(* IEC 61131-3 sources: TetherPLC/compat/tc2 (part 3) *)

(* ---- tc2_mc2_drive.st ---- *)
// tc2_mc2_drive.st — Tc2_MC2_Drive compatibility surface.
//
// TwinCAT's MC2 drive library addresses drives through AXIS_REF
// (here the flattened FB_MotionAxis UDINT handle, same convention
// as tc2_mc2.st).  Two transport families are covered:
//
//   CoE / OD  — CiA-402 object dictionary access through
//               FB_MotionAxis OP4/OP5 (works on both the in-process
//               tplc-motion backend and the Tether IO backend).
//               Manufacturer-specific sim objects 0x2002..0x2009
//               carry position offset, brake/park/CoE commands and
//               flying-saw characteristics (stored state, no
//               physical effect — documented).
//   SoE       — Sercos-over-EtherCAT mailbox through the builtin
//               FB_Soe (tplc-soe service, Tether IO only).  The
//               AXIS_REF handle maps to the SoE port as slave =
//               handle - 1 (MotionIoService assigns handle =
//               slave + 1).  In-process there is no SoE service,
//               so SoE FBs report bError/nErrorId = 99.
//
// NAME COLLISION NOTE: the SoE/AX5000 FB names match
// compat/tc2/tc2_drive.st (TwinCAT uses the same names in both
// libraries, differing only in the drive reference type).  This
// dialect has no library namespaces — link tc2_mc2_drive.st OR
// tc2_drive.st into a program, not both.
//
// Mapping notes (documented deviations):
//   - E_* enums (E_ParkMode, E_BrakeMode, E_PositionOffsetFeedback,
//     E_PositionOffsetMemory, E_DriveParameterNumber,
//     E_ReadWriteMode) are flattened to UDINT/INT inputs; values
//     are passed through to the backing object or ignored where
//     the sim has no equivalent.
//   - PVOID/ANY buffers (FB_CoERead/Write, FB_WriteDriveParameter)
//     are flattened to a single DINT Value; sub-index and
//     CompleteAccess are accepted but only sub-index 0 scalar
//     access is modeled.
//   - T_AmsNetID inputs are accepted for signature fidelity and
//     ignored (the axis reference already selects the drive).
//   - The 0x2002..0x2009 objects are stored command/state, not
//     physical: position offset is recorded but not applied to
//     motion, brake/park/CoE commands are recorded, saw
//     characteristics are read/write storage.
//
// SPDX-License-Identifier: Apache-2.0 OR MPL-2.0

// ---- shared helpers ------------------------------------------------
// SoE slave resolution: AXIS_REF handle -> SoE port address.
// (inlined per FB; handle = slave + 1 on the Tether IO backend)

// ================================================================== //
// §4.1 General Beckhoff
// ================================================================== //

// FB_ReadDriveParameter — read a drive parameter (OD object).
// ParameterNumber is the CiA402 object index; Mode 0 = single shot
// on Execute edge, Mode 1 = cyclic re-read while Execute is held
// (Interval is accepted; the scan rate is the cycle).
FUNCTION_BLOCK FB_ReadDriveParameter
VAR_INPUT
    Execute : BOOL;
    ParameterNumber : UDINT;
    Mode : UDINT;
    Interval : UDINT;
    Axis : UDINT;
END_VAR
VAR_OUTPUT
    Valid : BOOL;
    Value : DINT;
    Busy : BOOL;
    Done : BOOL;
    Error : BOOL;
    ErrorID : UDINT;
END_VAR
VAR
    ax : FB_MotionAxis;
    exPrev : BOOL;
    exEdge : BOOL;
END_VAR
    ax.AXIS := Axis;
    exEdge := Execute AND NOT exPrev; exPrev := Execute;
    Valid := FALSE; Busy := FALSE; Done := FALSE;
    Error := FALSE; ErrorID := 0;
    IF exEdge OR (Mode = 1 AND Execute) THEN
        ax.OP := 4;
        ax.INDEX := UDINT_TO_DINT(ParameterNumber);
        ax();
        IF ax.STATUS = 0 THEN
            Value := ax.VALUE;
            Valid := TRUE;
            IF exEdge THEN Done := TRUE; END_IF;
        ELSE
            Error := TRUE; ErrorID := ax.ERRID;
        END_IF;
    END_IF;
END_FUNCTION_BLOCK

// FB_WriteDriveParameter — write a drive parameter (OD object).
// Value is the flattened ANY buffer (single i32).
FUNCTION_BLOCK FB_WriteDriveParameter
VAR_INPUT
    Execute : BOOL;
    ParameterNumber : UDINT;
    Mode : UDINT;
    Interval : UDINT;
    Value : DINT;
    Axis : UDINT;
END_VAR
VAR_OUTPUT
    Valid : BOOL;
    Busy : BOOL;
    Done : BOOL;
    Error : BOOL;
    ErrorID : UDINT;
END_VAR
VAR
    ax : FB_MotionAxis;
    exPrev : BOOL;
    exEdge : BOOL;
END_VAR
    ax.AXIS := Axis;
    exEdge := Execute AND NOT exPrev; exPrev := Execute;
    Valid := FALSE; Busy := FALSE; Done := FALSE;
    Error := FALSE; ErrorID := 0;
    IF exEdge THEN
        ax.OP := 5;
        ax.INDEX := UDINT_TO_DINT(ParameterNumber);
        ax.VALUE := Value;
        ax();
        IF ax.STATUS = 0 THEN
            Valid := TRUE;
            Done := TRUE;
        ELSE
            Error := TRUE; ErrorID := ax.ERRID;
        END_IF;
    END_IF;
END_FUNCTION_BLOCK

// FB_SetPositionOffset — store a position offset (OD 0x2002).
// Absolute mode: offset = Position - PositionActualValue.
// Relative mode: offset accumulates (old + Position).  Feedback
// and Memory select encoder/drive/nameplate in TwinCAT; the sim
// has a single offset object, both are accepted and ignored.
FUNCTION_BLOCK FB_SetPositionOffset
VAR_INPUT
    Execute : BOOL;
    Position : LREAL;
    Relative : BOOL;
    Feedback : UDINT;
    Memory : UDINT;
    Axis : UDINT;
END_VAR
VAR_OUTPUT
    Busy : BOOL;
    Done : BOOL;
    Error : BOOL;
    ErrorID : UDINT;
END_VAR
VAR
    ax : FB_MotionAxis;
    exPrev : BOOL;
    exEdge : BOOL;
    posAct : DINT;
    offCur : DINT;
    np : DINT;
    p : DINT;
END_VAR
    ax.AXIS := Axis;
    exEdge := Execute AND NOT exPrev; exPrev := Execute;
    Busy := FALSE; Done := FALSE; Error := FALSE; ErrorID := 0;
    IF exEdge THEN
        p := LREAL_TO_DINT(Position);
        IF Relative THEN
            ax.OP := 4; ax.INDEX := 16#2002; ax();
            offCur := ax.VALUE;
            np := offCur + p;
        ELSE
            ax.OP := 4; ax.INDEX := 16#6064; ax();
            posAct := ax.VALUE;
            np := p - posAct;
        END_IF;
        ax.OP := 5; ax.INDEX := 16#2002; ax.VALUE := np; ax();
        IF ax.STATUS = 0 THEN
            Done := TRUE;
        ELSE
            Error := TRUE; ErrorID := ax.ERRID;
        END_IF;
    END_IF;
END_FUNCTION_BLOCK

// FB_DeletePositionOffset — clear the position offset (OD 0x2002).
FUNCTION_BLOCK FB_DeletePositionOffset
VAR_INPUT
    Execute : BOOL;
    Feedback : UDINT;
    Memory : UDINT;
    Axis : UDINT;
END_VAR
VAR_OUTPUT
    Busy : BOOL;
    Done : BOOL;
    Error : BOOL;
    ErrorID : UDINT;
END_VAR
VAR
    ax : FB_MotionAxis;
    exPrev : BOOL;
    exEdge : BOOL;
END_VAR
    ax.AXIS := Axis;
    exEdge := Execute AND NOT exPrev; exPrev := Execute;
    Busy := FALSE; Done := FALSE; Error := FALSE; ErrorID := 0;
    IF exEdge THEN
        ax.OP := 5; ax.INDEX := 16#2002; ax.VALUE := 0; ax();
        IF ax.STATUS = 0 THEN
            Done := TRUE;
        ELSE
            Error := TRUE; ErrorID := ax.ERRID;
        END_IF;
    END_IF;
END_FUNCTION_BLOCK

// FB_BrakeControl — brake command (OD 0x2003).  Mode is stored
// raw; the sim records the command without physical effect.
FUNCTION_BLOCK FB_BrakeControl
VAR_INPUT
    Execute : BOOL;
    Mode : UDINT;
    Axis : UDINT;
END_VAR
VAR_OUTPUT
    Busy : BOOL;
    Done : BOOL;
    Error : BOOL;
    ErrorID : UDINT;
END_VAR
VAR
    ax : FB_MotionAxis;
    exPrev : BOOL;
    exEdge : BOOL;
END_VAR
    ax.AXIS := Axis;
    exEdge := Execute AND NOT exPrev; exPrev := Execute;
    Busy := FALSE; Done := FALSE; Error := FALSE; ErrorID := 0;
    IF exEdge THEN
        ax.OP := 5; ax.INDEX := 16#2003;
        ax.VALUE := UDINT_TO_DINT(Mode); ax();
        IF ax.STATUS = 0 THEN
            Done := TRUE;
        ELSE
            Error := TRUE; ErrorID := ax.ERRID;
        END_IF;
    END_IF;
END_FUNCTION_BLOCK

// FB_ParkAxis — park/release via the SoE park mailbox (OP 7).
// Mode 0 = release, nonzero = park.  Requires the SoE backend
// (Tether IO); in-process reports bError.
FUNCTION_BLOCK FB_ParkAxis
VAR_INPUT
    Execute : BOOL;
    Mode : UDINT;
    NetId : STRING[15];
    Axis : UDINT;
END_VAR
VAR_OUTPUT
    Busy : BOOL;
    Done : BOOL;
    Error : BOOL;
    ErrorID : UDINT;
END_VAR
VAR
    raw : FB_Soe;
    exPrev : BOOL;
    exEdge : BOOL;
    slave : UDINT;
END_VAR
    exEdge := Execute AND NOT exPrev; exPrev := Execute;
    IF Axis > 0 THEN slave := Axis - 1; ELSE slave := 0; END_IF;
    Busy := FALSE; Done := FALSE; Error := FALSE; ErrorID := 0;
    IF exEdge THEN
        raw.OP := 7;
        raw.SLAVE := slave;
        IF Mode <> 0 THEN raw.VALUE := 1; ELSE raw.VALUE := 0; END_IF;
        raw();
        IF raw.STATUS < 0 THEN
            Error := TRUE; ErrorID := raw.ERRID;
        ELSE
            Done := TRUE;
        END_IF;
    END_IF;
END_FUNCTION_BLOCK

// FB_ReadDriveInfo — axis/drive info snapshot (FB_MotionAxis OP6).
FUNCTION_BLOCK FB_ReadDriveInfo
VAR_INPUT
    Execute : BOOL;
    Axis : UDINT;
END_VAR
VAR_OUTPUT
    Valid : BOOL;
    State : DINT;
    Fault : DINT;
    ModeOp : DINT;
    TargetReached : BOOL;
    PosActual : DINT;
    VelActual : DINT;
    Busy : BOOL;
    Done : BOOL;
    Error : BOOL;
    ErrorID : UDINT;
END_VAR
VAR
    ax : FB_MotionAxis;
    exPrev : BOOL;
    exEdge : BOOL;
END_VAR
    ax.AXIS := Axis;
    exEdge := Execute AND NOT exPrev; exPrev := Execute;
    Valid := FALSE; Busy := FALSE; Done := FALSE;
    Error := FALSE; ErrorID := 0;
    IF exEdge THEN
        ax.OP := 6; ax();
        IF ax.STATUS < 0 THEN
            Error := TRUE; ErrorID := ax.ERRID;
        ELSE
            Valid := TRUE;
            Done := TRUE;
            State := ax.STATUS;
            Fault := ax.FAULT;
            ModeOp := ax.MODE;
            TargetReached := (ax.TARGET_REACHED <> 0);
            PosActual := ax.POS_ACTUAL;
            VelActual := ax.VEL_ACTUAL;
        END_IF;
    END_IF;
END_FUNCTION_BLOCK

// ================================================================== //
// §4.2 General SoE
// ================================================================== //
// All SoE FBs resolve slave = Axis - 1 and drive the FB_Soe builtin.

// FB_SoERead — generic SoE element read.  Index is the SoE element
// id; the supported subset is the state-snapshot fields:
//   16#0135 -> status word (S-0-0135), 16#0267 -> password.
// Other element ids report Error (arbitrary P-0-xxxx access is not
// modeled).  Value is LREAL; u16/u32 fields are returned raw.
FUNCTION_BLOCK FB_SoERead
VAR_INPUT
    Execute : BOOL;
    Index : UDINT;
    NetId : STRING[15];
    Axis : UDINT;
END_VAR
VAR_OUTPUT
    Value : LREAL;
    Busy : BOOL;
    Done : BOOL;
    Error : BOOL;
    ErrorID : UDINT;
END_VAR
VAR
    raw : FB_Soe;
    exPrev : BOOL;
    exEdge : BOOL;
    slave : UDINT;
END_VAR
    exEdge := Execute AND NOT exPrev; exPrev := Execute;
    IF Axis > 0 THEN slave := Axis - 1; ELSE slave := 0; END_IF;
    Busy := FALSE; Done := FALSE; Error := FALSE; ErrorID := 0;
    IF exEdge THEN
        raw.OP := 1;
        raw.SLAVE := slave;
        raw();
        IF raw.STATUS < 0 THEN
            Error := TRUE; ErrorID := raw.ERRID;
        ELSE
            IF Index = 16#0135 THEN
                Value := UDINT_TO_LREAL(raw.STATUSW);
                Done := TRUE;
            ELSIF Index = 16#0267 THEN
                Value := UDINT_TO_LREAL(raw.PASSWD);
                Done := TRUE;
            ELSE
                Error := TRUE; ErrorID := 2;
            END_IF;
        END_IF;
    END_IF;
END_FUNCTION_BLOCK

// FB_SoEWrite — generic SoE element write.  Supported subset:
// Index 16#0267 -> drive password (S-0-0267).  Other ids report
// Error (arbitrary P-0-xxxx writes are not modeled).
FUNCTION_BLOCK FB_SoEWrite
VAR_INPUT
    Execute : BOOL;
    Index : UDINT;
    Value : DINT;
    NetId : STRING[15];
    Axis : UDINT;
END_VAR
VAR_OUTPUT
    Busy : BOOL;
    Done : BOOL;
    Error : BOOL;
    ErrorID : UDINT;
END_VAR
VAR
    raw : FB_Soe;
    exPrev : BOOL;
    exEdge : BOOL;
    slave : UDINT;
END_VAR
    exEdge := Execute AND NOT exPrev; exPrev := Execute;
    IF Axis > 0 THEN slave := Axis - 1; ELSE slave := 0; END_IF;
    Busy := FALSE; Done := FALSE; Error := FALSE; ErrorID := 0;
    IF exEdge THEN
        IF Index = 16#0267 THEN
            raw.OP := 2;
            raw.SLAVE := slave;
            raw.VALUE := Value;
            raw();
            IF raw.STATUS < 0 THEN
                Error := TRUE; ErrorID := raw.ERRID;
            ELSE
                Done := TRUE;
            END_IF;
        ELSE
            Error := TRUE; ErrorID := 2;
        END_IF;
    END_IF;
END_FUNCTION_BLOCK

// FB_SoESetDataAccessMode — SoE parameter access mode.  The sim
// mailbox always uses parallel access; the FB accepts the request
// and completes (documented no-op).
FUNCTION_BLOCK FB_SoESetDataAccessMode
VAR_INPUT
    Execute : BOOL;
    Mode : UDINT;
    Axis : UDINT;
END_VAR
VAR_OUTPUT
    Busy : BOOL;
    Done : BOOL;
    Error : BOOL;
    ErrorID : UDINT;
END_VAR
VAR
    exPrev : BOOL;
    exEdge : BOOL;
END_VAR
    exEdge := Execute AND NOT exPrev; exPrev := Execute;
    Busy := FALSE; Done := FALSE; Error := FALSE; ErrorID := 0;
    IF exEdge THEN
        Done := TRUE;
    END_IF;
END_FUNCTION_BLOCK

// ---- command FBs ----------------------------------------------------

// FB_SoEReset — S-0-0099 drive reset.
FUNCTION_BLOCK FB_SoEReset
VAR_INPUT
    Execute : BOOL;
    NetId : STRING[15];
    Axis : UDINT;
END_VAR
VAR_OUTPUT
    Busy : BOOL;
    Done : BOOL;
    Error : BOOL;
    ErrorID : UDINT;
END_VAR
VAR
    raw : FB_Soe;
    exPrev : BOOL;
    exEdge : BOOL;
    slave : UDINT;
END_VAR
    exEdge := Execute AND NOT exPrev; exPrev := Execute;
    IF Axis > 0 THEN slave := Axis - 1; ELSE slave := 0; END_IF;
    Busy := FALSE; Done := FALSE; Error := FALSE; ErrorID := 0;
    IF exEdge THEN
        raw.OP := 5;
        raw.SLAVE := slave;
        raw();
        IF raw.STATUS < 0 THEN
            Error := TRUE; ErrorID := raw.ERRID;
        ELSE
            Done := TRUE;
        END_IF;
    END_IF;
END_FUNCTION_BLOCK

// FB_SoEWritePassword — S-0-0267 drive password.
FUNCTION_BLOCK FB_SoEWritePassword
VAR_INPUT
    Execute : BOOL;
    Password : UDINT;
    NetId : STRING[15];
    Axis : UDINT;
END_VAR
VAR_OUTPUT
    Busy : BOOL;
    Done : BOOL;
    Error : BOOL;
    ErrorID : UDINT;
END_VAR
VAR
    raw : FB_Soe;
    exPrev : BOOL;
    exEdge : BOOL;
    slave : UDINT;
END_VAR
    exEdge := Execute AND NOT exPrev; exPrev := Execute;
    IF Axis > 0 THEN slave := Axis - 1; ELSE slave := 0; END_IF;
    Busy := FALSE; Done := FALSE; Error := FALSE; ErrorID := 0;
    IF exEdge THEN
        raw.OP := 2;
        raw.SLAVE := slave;
        raw.VALUE := UDINT_TO_DINT(Password);
        raw();
        IF raw.STATUS < 0 THEN
            Error := TRUE; ErrorID := raw.ERRID;
        ELSE
            Done := TRUE;
        END_IF;
    END_IF;
END_FUNCTION_BLOCK

// FB_SoEExecuteCommand — execute an SoE command id.
FUNCTION_BLOCK FB_SoEExecuteCommand
VAR_INPUT
    Execute : BOOL;
    CommandId : UDINT;
    NetId : STRING[15];
    Axis : UDINT;
END_VAR
VAR_OUTPUT
    Busy : BOOL;
    Done : BOOL;
    Error : BOOL;
    ErrorID : UDINT;
END_VAR
VAR
    raw : FB_Soe;
    exPrev : BOOL;
    exEdge : BOOL;
    slave : UDINT;
END_VAR
    exEdge := Execute AND NOT exPrev; exPrev := Execute;
    IF Axis > 0 THEN slave := Axis - 1; ELSE slave := 0; END_IF;
    Busy := FALSE; Done := FALSE; Error := FALSE; ErrorID := 0;
    IF exEdge THEN
        raw.OP := 4;
        raw.SLAVE := slave;
        raw.VALUE := UDINT_TO_DINT(CommandId);
        raw();
        IF raw.STATUS < 0 THEN
            Error := TRUE; ErrorID := raw.ERRID;
        ELSE
            Done := TRUE;
        END_IF;
    END_IF;
END_FUNCTION_BLOCK

// FB_SoEWriteCommandControl — command control word.
FUNCTION_BLOCK FB_SoEWriteCommandControl
VAR_INPUT
    Execute : BOOL;
    CommandControl : UDINT;
    NetId : STRING[15];
    Axis : UDINT;
END_VAR
VAR_OUTPUT
    Busy : BOOL;
    Done : BOOL;
    Error : BOOL;
    ErrorID : UDINT;
END_VAR
VAR
    raw : FB_Soe;
    exPrev : BOOL;
    exEdge : BOOL;
    slave : UDINT;
END_VAR
    exEdge := Execute AND NOT exPrev; exPrev := Execute;
    IF Axis > 0 THEN slave := Axis - 1; ELSE slave := 0; END_IF;
    Busy := FALSE; Done := FALSE; Error := FALSE; ErrorID := 0;
    IF exEdge THEN
        raw.OP := 3;
        raw.SLAVE := slave;
        raw.VALUE := UDINT_TO_DINT(CommandControl);
        raw();
        IF raw.STATUS < 0 THEN
            Error := TRUE; ErrorID := raw.ERRID;
        ELSE
            Done := TRUE;
        END_IF;
    END_IF;
END_FUNCTION_BLOCK

// FB_SoEReadCommandState — SoE command state
// (0 idle, 1 running, 2 done, 3 error).
FUNCTION_BLOCK FB_SoEReadCommandState
VAR_INPUT
    Execute : BOOL;
    NetId : STRING[15];
    Axis : UDINT;
END_VAR
VAR_OUTPUT
    CommandState : UDINT;
    Busy : BOOL;
    Done : BOOL;
    Error : BOOL;
    ErrorID : UDINT;
END_VAR
VAR
    raw : FB_Soe;
    exPrev : BOOL;
    exEdge : BOOL;
    slave : UDINT;
END_VAR
    exEdge := Execute AND NOT exPrev; exPrev := Execute;
    IF Axis > 0 THEN slave := Axis - 1; ELSE slave := 0; END_IF;
    Busy := FALSE; Done := FALSE; Error := FALSE; ErrorID := 0;
    IF exEdge THEN
        raw.OP := 1;
        raw.SLAVE := slave;
        raw();
        IF raw.STATUS < 0 THEN
            Error := TRUE; ErrorID := raw.ERRID;
        ELSE
            CommandState := raw.CMDSTATE;
            Done := TRUE;
        END_IF;
    END_IF;
END_FUNCTION_BLOCK

// ---- diagnostics FBs -------------------------------------------------

// FB_SoEReadDiagMessage — S-0-0095 diagnosis message.
FUNCTION_BLOCK FB_SoEReadDiagMessage
VAR_INPUT
    Execute : BOOL;
    NetId : STRING[15];
    Axis : UDINT;
END_VAR
VAR_OUTPUT
    DiagMessage : STRING[63];
    Busy : BOOL;
    Done : BOOL;
    Error : BOOL;
    ErrorID : UDINT;
END_VAR
VAR
    raw : FB_Soe;
    exPrev : BOOL;
    exEdge : BOOL;
    slave : UDINT;
END_VAR
    exEdge := Execute AND NOT exPrev; exPrev := Execute;
    IF Axis > 0 THEN slave := Axis - 1; ELSE slave := 0; END_IF;
    Busy := FALSE; Done := FALSE; Error := FALSE; ErrorID := 0;
    IF exEdge THEN
        raw.OP := 1;
        raw.SLAVE := slave;
        raw();
        IF raw.STATUS < 0 THEN
            Error := TRUE; ErrorID := raw.ERRID;
        ELSE
            DiagMessage := raw.DIAGMSG;
            Done := TRUE;
        END_IF;
    END_IF;
END_FUNCTION_BLOCK

// FB_SoEReadDiagNumber — diagnosis number.
FUNCTION_BLOCK FB_SoEReadDiagNumber
VAR_INPUT
    Execute : BOOL;
    NetId : STRING[15];
    Axis : UDINT;
END_VAR
VAR_OUTPUT
    DiagNumber : UDINT;
    Busy : BOOL;
    Done : BOOL;
    Error : BOOL;
    ErrorID : UDINT;
END_VAR
VAR
    raw : FB_Soe;
    exPrev : BOOL;
    exEdge : BOOL;
    slave : UDINT;
END_VAR
    exEdge := Execute AND NOT exPrev; exPrev := Execute;
    IF Axis > 0 THEN slave := Axis - 1; ELSE slave := 0; END_IF;
    Busy := FALSE; Done := FALSE; Error := FALSE; ErrorID := 0;
    IF exEdge THEN
        raw.OP := 1;
        raw.SLAVE := slave;
        raw();
        IF raw.STATUS < 0 THEN
            Error := TRUE; ErrorID := raw.ERRID;
        ELSE
            DiagNumber := raw.DIAGNUM;
            Done := TRUE;
        END_IF;
    END_IF;
END_FUNCTION_BLOCK

// FB_SoEReadDiagNumberList — diagnosis number list (flattened:
// DiagCount + DiagList internal array).
FUNCTION_BLOCK FB_SoEReadDiagNumberList
VAR_INPUT
    Execute : BOOL;
    NetId : STRING[15];
    Axis : UDINT;
END_VAR
VAR_OUTPUT
    DiagCount : UDINT;
    Busy : BOOL;
    Done : BOOL;
    Error : BOOL;
    ErrorID : UDINT;
END_VAR
VAR
    raw : FB_Soe;
    exPrev : BOOL;
    exEdge : BOOL;
    slave : UDINT;
    i : UDINT;
    DiagList : ARRAY[0..7] OF UDINT;
END_VAR
    exEdge := Execute AND NOT exPrev; exPrev := Execute;
    IF Axis > 0 THEN slave := Axis - 1; ELSE slave := 0; END_IF;
    Busy := FALSE; Done := FALSE; Error := FALSE; ErrorID := 0;
    IF exEdge THEN
        raw.OP := 1;
        raw.SLAVE := slave;
        raw();
        IF raw.STATUS < 0 THEN
            Error := TRUE; ErrorID := raw.ERRID;
        ELSE
            DiagCount := raw.DIAGCOUNT;
            FOR i := 0 TO 7 DO
                DiagList[i] := raw.DIAGLIST[i];
            END_FOR;
            Done := TRUE;
        END_IF;
    END_IF;
END_FUNCTION_BLOCK

// FB_SoEReadClassXDiag — class-X diagnosis.
FUNCTION_BLOCK FB_SoEReadClassXDiag
VAR_INPUT
    Execute : BOOL;
    NetId : STRING[15];
    Axis : UDINT;
END_VAR
VAR_OUTPUT
    ClassXDiag : UDINT;
    Busy : BOOL;
    Done : BOOL;
    Error : BOOL;
    ErrorID : UDINT;
END_VAR
VAR
    raw : FB_Soe;
    exPrev : BOOL;
    exEdge : BOOL;
    slave : UDINT;
END_VAR
    exEdge := Execute AND NOT exPrev; exPrev := Execute;
    IF Axis > 0 THEN slave := Axis - 1; ELSE slave := 0; END_IF;
    Busy := FALSE; Done := FALSE; Error := FALSE; ErrorID := 0;
    IF exEdge THEN
        raw.OP := 1;
        raw.SLAVE := slave;
        raw();
        IF raw.STATUS < 0 THEN
            Error := TRUE; ErrorID := raw.ERRID;
        ELSE
            ClassXDiag := raw.CLASSX;
            Done := TRUE;
        END_IF;
    END_IF;
END_FUNCTION_BLOCK

// ---- current-value readers -------------------------------------------

FUNCTION_BLOCK FB_SoEReadAmplifierTemperature
VAR_INPUT
    Execute : BOOL;
    NetId : STRING[15];
    Axis : UDINT;
END_VAR
VAR_OUTPUT
    Value : LREAL;
    Busy : BOOL;
    Done : BOOL;
    Error : BOOL;
    ErrorID : UDINT;
END_VAR
VAR
    raw : FB_Soe;
    exPrev : BOOL;
    exEdge : BOOL;
    slave : UDINT;
END_VAR
    exEdge := Execute AND NOT exPrev; exPrev := Execute;
    IF Axis > 0 THEN slave := Axis - 1; ELSE slave := 0; END_IF;
    Busy := FALSE; Done := FALSE; Error := FALSE; ErrorID := 0;
    IF exEdge THEN
        raw.OP := 1;
        raw.SLAVE := slave;
        raw();
        IF raw.STATUS < 0 THEN
            Error := TRUE; ErrorID := raw.ERRID;
        ELSE
            Value := raw.AMPTEMP;
            Done := TRUE;
        END_IF;
    END_IF;
END_FUNCTION_BLOCK

FUNCTION_BLOCK FB_SoEReadMotorTemperature
VAR_INPUT
    Execute : BOOL;
    NetId : STRING[15];
    Axis : UDINT;
END_VAR
VAR_OUTPUT
    Value : LREAL;
    Busy : BOOL;
    Done : BOOL;
    Error : BOOL;
    ErrorID : UDINT;
END_VAR
VAR
    raw : FB_Soe;
    exPrev : BOOL;
    exEdge : BOOL;
    slave : UDINT;
END_VAR
    exEdge := Execute AND NOT exPrev; exPrev := Execute;
    IF Axis > 0 THEN slave := Axis - 1; ELSE slave := 0; END_IF;
    Busy := FALSE; Done := FALSE; Error := FALSE; ErrorID := 0;
    IF exEdge THEN
        raw.OP := 1;
        raw.SLAVE := slave;
        raw();
        IF raw.STATUS < 0 THEN
            Error := TRUE; ErrorID := raw.ERRID;
        ELSE
            Value := raw.MTEMPT;
            Done := TRUE;
        END_IF;
    END_IF;
END_FUNCTION_BLOCK

FUNCTION_BLOCK FB_SoEReadDcBusVoltage
VAR_INPUT
    Execute : BOOL;
    NetId : STRING[15];
    Axis : UDINT;
END_VAR
VAR_OUTPUT
    Value : LREAL;
    Busy : BOOL;
    Done : BOOL;
    Error : BOOL;
    ErrorID : UDINT;
END_VAR
VAR
    raw : FB_Soe;
    exPrev : BOOL;
    exEdge : BOOL;
    slave : UDINT;
END_VAR
    exEdge := Execute AND NOT exPrev; exPrev := Execute;
    IF Axis > 0 THEN slave := Axis - 1; ELSE slave := 0; END_IF;
    Busy := FALSE; Done := FALSE; Error := FALSE; ErrorID := 0;
    IF exEdge THEN
        raw.OP := 1;
        raw.SLAVE := slave;
        raw();
        IF raw.STATUS < 0 THEN
            Error := TRUE; ErrorID := raw.ERRID;
        ELSE
            Value := raw.DCVOLT;
            Done := TRUE;
        END_IF;
    END_IF;
END_FUNCTION_BLOCK

FUNCTION_BLOCK FB_SoEReadDcBusCurrent
VAR_INPUT
    Execute : BOOL;
    NetId : STRING[15];
    Axis : UDINT;
END_VAR
VAR_OUTPUT
    Value : LREAL;
    Busy : BOOL;
    Done : BOOL;
    Error : BOOL;
    ErrorID : UDINT;
END_VAR
VAR
    raw : FB_Soe;
    exPrev : BOOL;
    exEdge : BOOL;
    slave : UDINT;
END_VAR
    exEdge := Execute AND NOT exPrev; exPrev := Execute;
    IF Axis > 0 THEN slave := Axis - 1; ELSE slave := 0; END_IF;
    Busy := FALSE; Done := FALSE; Error := FALSE; ErrorID := 0;
    IF exEdge THEN
        raw.OP := 1;
        raw.SLAVE := slave;
        raw();
        IF raw.STATUS < 0 THEN
            Error := TRUE; ErrorID := raw.ERRID;
        ELSE
            Value := raw.DCCURR;
            Done := TRUE;
        END_IF;
    END_IF;
END_FUNCTION_BLOCK

// ================================================================== //
// §4.3 General CoE — SDO object access via FB_MotionAxis OP4/OP5.
// Index/SubIndex select the object; SubIndex and CompleteAccess are
// accepted but only sub-index 0 scalar access is modeled.  Value is
// the flattened PVOID buffer (single i32).
// ================================================================== //

// FB_CoERead — CoE SDO upload.
FUNCTION_BLOCK FB_CoERead
VAR_INPUT
    Execute : BOOL;
    Index : UDINT;
    SubIndex : UDINT;
    CompleteAccess : BOOL;
    NetId : STRING[15];
    Axis : UDINT;
END_VAR
VAR_OUTPUT
    Value : DINT;
    Busy : BOOL;
    Done : BOOL;
    Error : BOOL;
    ErrorID : UDINT;
END_VAR
VAR
    ax : FB_MotionAxis;
    exPrev : BOOL;
    exEdge : BOOL;
END_VAR
    ax.AXIS := Axis;
    exEdge := Execute AND NOT exPrev; exPrev := Execute;
    Busy := FALSE; Done := FALSE; Error := FALSE; ErrorID := 0;
    IF exEdge THEN
        IF SubIndex <> 0 THEN
            Error := TRUE; ErrorID := 2;   // sub-index unsupported
        ELSE
            ax.OP := 4;
            ax.INDEX := UDINT_TO_DINT(Index);
            ax();
            IF ax.STATUS = 0 THEN
                Value := ax.VALUE;
                Done := TRUE;
            ELSE
                Error := TRUE; ErrorID := ax.ERRID;
            END_IF;
        END_IF;
    END_IF;
END_FUNCTION_BLOCK

// FB_CoEWrite — CoE SDO download.
FUNCTION_BLOCK FB_CoEWrite
VAR_INPUT
    Execute : BOOL;
    Index : UDINT;
    SubIndex : UDINT;
    Value : DINT;
    CompleteAccess : BOOL;
    NetId : STRING[15];
    Axis : UDINT;
END_VAR
VAR_OUTPUT
    Busy : BOOL;
    Done : BOOL;
    Error : BOOL;
    ErrorID : UDINT;
END_VAR
VAR
    ax : FB_MotionAxis;
    exPrev : BOOL;
    exEdge : BOOL;
END_VAR
    ax.AXIS := Axis;
    exEdge := Execute AND NOT exPrev; exPrev := Execute;
    Busy := FALSE; Done := FALSE; Error := FALSE; ErrorID := 0;
    IF exEdge THEN
        IF SubIndex <> 0 THEN
            Error := TRUE; ErrorID := 2;
        ELSE
            ax.OP := 5;
            ax.INDEX := UDINT_TO_DINT(Index);
            ax.VALUE := Value;
            ax();
            IF ax.STATUS = 0 THEN
                Done := TRUE;
            ELSE
                Error := TRUE; ErrorID := ax.ERRID;
            END_IF;
        END_IF;
    END_IF;
END_FUNCTION_BLOCK

// FB_CoEExecuteCommand — execute a CoE drive command (OD 0x2005).
// Command is the flattened command id; the sim records it.
FUNCTION_BLOCK FB_CoEExecuteCommand
VAR_INPUT
    Execute : BOOL;
    Command : UDINT;
    NetId : STRING[15];
    Axis : UDINT;
END_VAR
VAR_OUTPUT
    Busy : BOOL;
    Done : BOOL;
    Error : BOOL;
    ErrorID : UDINT;
END_VAR
VAR
    ax : FB_MotionAxis;
    exPrev : BOOL;
    exEdge : BOOL;
END_VAR
    ax.AXIS := Axis;
    exEdge := Execute AND NOT exPrev; exPrev := Execute;
    Busy := FALSE; Done := FALSE; Error := FALSE; ErrorID := 0;
    IF exEdge THEN
        ax.OP := 5; ax.INDEX := 16#2005;
        ax.VALUE := UDINT_TO_DINT(Command); ax();
        IF ax.STATUS = 0 THEN
            Done := TRUE;
        ELSE
            Error := TRUE; ErrorID := ax.ERRID;
        END_IF;
    END_IF;
END_FUNCTION_BLOCK

// ================================================================== //
// §4.4 AX5000 SoE — same SoE mailbox surface as the general blocks,
// AX5000-specific objects (mains voltage, motor ctrl word, firmware,
// park, position offset).
// ================================================================== //

// FB_SoEAX5000ReadActMainVoltage — P-0-0200 peak mains voltage.
FUNCTION_BLOCK FB_SoEAX5000ReadActMainVoltage
VAR_INPUT
    Execute : BOOL;
    NetId : STRING[15];
    Axis : UDINT;
END_VAR
VAR_OUTPUT
    Voltage : LREAL;
    Busy : BOOL;
    Done : BOOL;
    Error : BOOL;
    ErrorID : UDINT;
END_VAR
VAR
    raw : FB_Soe;
    exPrev : BOOL;
    exEdge : BOOL;
    slave : UDINT;
END_VAR
    exEdge := Execute AND NOT exPrev; exPrev := Execute;
    IF Axis > 0 THEN slave := Axis - 1; ELSE slave := 0; END_IF;
    Busy := FALSE; Done := FALSE; Error := FALSE; ErrorID := 0;
    IF exEdge THEN
        raw.OP := 1;
        raw.SLAVE := slave;
        raw();
        IF raw.STATUS < 0 THEN
            Error := TRUE; ErrorID := raw.ERRID;
        ELSE
            Voltage := raw.AXMAINS;
            Done := TRUE;
        END_IF;
    END_IF;
END_FUNCTION_BLOCK

// FB_SoEAX5000SetMotorCtrlWord — motor control word (mailbox OP6).
// bForceUnlock accepted for signature compatibility.
FUNCTION_BLOCK FB_SoEAX5000SetMotorCtrlWord
VAR_INPUT
    Execute : BOOL;
    MotorCtrlWord : UDINT;
    bForceUnlock : BOOL;
    NetId : STRING[15];
    Axis : UDINT;
END_VAR
VAR_OUTPUT
    Busy : BOOL;
    Done : BOOL;
    Error : BOOL;
    ErrorID : UDINT;
END_VAR
VAR
    raw : FB_Soe;
    exPrev : BOOL;
    exEdge : BOOL;
    slave : UDINT;
END_VAR
    exEdge := Execute AND NOT exPrev; exPrev := Execute;
    IF Axis > 0 THEN slave := Axis - 1; ELSE slave := 0; END_IF;
    Busy := FALSE; Done := FALSE; Error := FALSE; ErrorID := 0;
    IF exEdge THEN
        raw.OP := 6;
        raw.SLAVE := slave;
        raw.VALUE := UDINT_TO_DINT(MotorCtrlWord);
        raw();
        IF raw.STATUS < 0 THEN
            Error := TRUE; ErrorID := raw.ERRID;
        ELSE
            Done := TRUE;
        END_IF;
    END_IF;
END_FUNCTION_BLOCK

// FB_SoEAX5000FirmwareUpdate — reports simulated firmware
// revision/build; no firmware pool or flashing is simulated.
FUNCTION_BLOCK FB_SoEAX5000FirmwareUpdate
VAR_INPUT
    Execute : BOOL;
    NetId : STRING[15];
    Axis : UDINT;
END_VAR
VAR_OUTPUT
    FirmwareRevision : UDINT;
    FirmwareBuild : UDINT;
    Busy : BOOL;
    Done : BOOL;
    Error : BOOL;
    ErrorID : UDINT;
END_VAR
VAR
    raw : FB_Soe;
    exPrev : BOOL;
    exEdge : BOOL;
    slave : UDINT;
END_VAR
    exEdge := Execute AND NOT exPrev; exPrev := Execute;
    IF Axis > 0 THEN slave := Axis - 1; ELSE slave := 0; END_IF;
    Busy := FALSE; Done := FALSE; Error := FALSE; ErrorID := 0;
    IF exEdge THEN
        raw.OP := 1;
        raw.SLAVE := slave;
        raw();
        IF raw.STATUS < 0 THEN
            Error := TRUE; ErrorID := raw.ERRID;
        ELSE
            FirmwareRevision := raw.AXFWREV;
            FirmwareBuild := raw.AXFWBUILD;
            Done := TRUE;
        END_IF;
    END_IF;
END_FUNCTION_BLOCK

// FB_SoEAX5000SetPositionOffset — AX5000 position offset (OD 0x2002).
FUNCTION_BLOCK FB_SoEAX5000SetPositionOffset
VAR_INPUT
    Execute : BOOL;
    Position : LREAL;
    Relative : BOOL;
    Feedback : UDINT;
    Memory : UDINT;
    NetId : STRING[15];
    Axis : UDINT;
END_VAR
VAR_OUTPUT
    Busy : BOOL;
    Done : BOOL;
    Error : BOOL;
    ErrorID : UDINT;
END_VAR
VAR
    ax : FB_MotionAxis;
    exPrev : BOOL;
    exEdge : BOOL;
    posAct : DINT;
    np : DINT;
    p : DINT;
END_VAR
    ax.AXIS := Axis;
    exEdge := Execute AND NOT exPrev; exPrev := Execute;
    Busy := FALSE; Done := FALSE; Error := FALSE; ErrorID := 0;
    IF exEdge THEN
        p := LREAL_TO_DINT(Position);
        IF Relative THEN
            np := p;                    // relative: offset delta
        ELSE
            ax.OP := 4; ax.INDEX := 16#6064; ax();
            posAct := ax.VALUE;
            np := p - posAct;
        END_IF;
        ax.OP := 5; ax.INDEX := 16#2002; ax.VALUE := np; ax();
        IF ax.STATUS = 0 THEN
            Done := TRUE;
        ELSE
            Error := TRUE; ErrorID := ax.ERRID;
        END_IF;
    END_IF;
END_FUNCTION_BLOCK

// FB_SoEAX5000DeletePositionOffset — clear AX5000 position offset.
FUNCTION_BLOCK FB_SoEAX5000DeletePositionOffset
VAR_INPUT
    Execute : BOOL;
    Feedback : UDINT;
    Memory : UDINT;
    NetId : STRING[15];
    Axis : UDINT;
END_VAR
VAR_OUTPUT
    Busy : BOOL;
    Done : BOOL;
    Error : BOOL;
    ErrorID : UDINT;
END_VAR
VAR
    ax : FB_MotionAxis;
    exPrev : BOOL;
    exEdge : BOOL;
END_VAR
    ax.AXIS := Axis;
    exEdge := Execute AND NOT exPrev; exPrev := Execute;
    Busy := FALSE; Done := FALSE; Error := FALSE; ErrorID := 0;
    IF exEdge THEN
        ax.OP := 5; ax.INDEX := 16#2002; ax.VALUE := 0; ax();
        IF ax.STATUS = 0 THEN
            Done := TRUE;
        ELSE
            Error := TRUE; ErrorID := ax.ERRID;
        END_IF;
    END_IF;
END_FUNCTION_BLOCK

// FB_SoEAX5000ParkAxis — park/unpark via SoE mailbox (OP 7).
FUNCTION_BLOCK FB_SoEAX5000ParkAxis
VAR_INPUT
    Execute : BOOL;
    Mode : UDINT;
    NetId : STRING[15];
    Axis : UDINT;
END_VAR
VAR_OUTPUT
    Busy : BOOL;
    Done : BOOL;
    Error : BOOL;
    ErrorID : UDINT;
END_VAR
VAR
    raw : FB_Soe;
    exPrev : BOOL;
    exEdge : BOOL;
    slave : UDINT;
END_VAR
    exEdge := Execute AND NOT exPrev; exPrev := Execute;
    IF Axis > 0 THEN slave := Axis - 1; ELSE slave := 0; END_IF;
    Busy := FALSE; Done := FALSE; Error := FALSE; ErrorID := 0;
    IF exEdge THEN
        raw.OP := 7;
        raw.SLAVE := slave;
        IF Mode <> 0 THEN raw.VALUE := 1; ELSE raw.VALUE := 0; END_IF;
        raw();
        IF raw.STATUS < 0 THEN
            Error := TRUE; ErrorID := raw.ERRID;
        ELSE
            Done := TRUE;
        END_IF;
    END_IF;
END_FUNCTION_BLOCK

// ================================================================== //
// §4.5 AX8000 CoE — brake/park/offset over OD objects 0x2002-0x2004.
// ================================================================== //

// FB_CoEAX8000BrakeControl — AX8000 brake (OD 0x2003).
FUNCTION_BLOCK FB_CoEAX8000BrakeControl
VAR_INPUT
    Execute : BOOL;
    Mode : UDINT;
    NetId : STRING[15];
    Axis : UDINT;
END_VAR
VAR_OUTPUT
    Busy : BOOL;
    Done : BOOL;
    Error : BOOL;
    ErrorID : UDINT;
END_VAR
VAR
    ax : FB_MotionAxis;
    exPrev : BOOL;
    exEdge : BOOL;
END_VAR
    ax.AXIS := Axis;
    exEdge := Execute AND NOT exPrev; exPrev := Execute;
    Busy := FALSE; Done := FALSE; Error := FALSE; ErrorID := 0;
    IF exEdge THEN
        ax.OP := 5; ax.INDEX := 16#2003;
        ax.VALUE := UDINT_TO_DINT(Mode); ax();
        IF ax.STATUS = 0 THEN
            Done := TRUE;
        ELSE
            Error := TRUE; ErrorID := ax.ERRID;
        END_IF;
    END_IF;
END_FUNCTION_BLOCK

// FB_CoEAX8000BrakeTest — brake test: writes the test command and
// reports Succeeded (the sim has no torque verification; the test
// always succeeds once the command is accepted — documented).
FUNCTION_BLOCK FB_CoEAX8000BrakeTest
VAR_INPUT
    Execute : BOOL;
    NetId : STRING[15];
    Axis : UDINT;
END_VAR
VAR_OUTPUT
    Succeeded : BOOL;
    Busy : BOOL;
    Done : BOOL;
    Error : BOOL;
    ErrorID : UDINT;
END_VAR
VAR
    ax : FB_MotionAxis;
    exPrev : BOOL;
    exEdge : BOOL;
END_VAR
    ax.AXIS := Axis;
    exEdge := Execute AND NOT exPrev; exPrev := Execute;
    Busy := FALSE; Done := FALSE; Error := FALSE; ErrorID := 0;
    Succeeded := FALSE;
    IF exEdge THEN
        ax.OP := 5; ax.INDEX := 16#2003; ax.VALUE := 2; ax();
        IF ax.STATUS = 0 THEN
            Done := TRUE;
            Succeeded := TRUE;
        ELSE
            Error := TRUE; ErrorID := ax.ERRID;
        END_IF;
    END_IF;
END_FUNCTION_BLOCK

// FB_CoEAX8000SetPositionOffset — AX8000 position offset (0x2002).
FUNCTION_BLOCK FB_CoEAX8000SetPositionOffset
VAR_INPUT
    Execute : BOOL;
    Position : LREAL;
    Relative : BOOL;
    Feedback : UDINT;
    Memory : UDINT;
    NetId : STRING[15];
    Axis : UDINT;
END_VAR
VAR_OUTPUT
    Busy : BOOL;
    Done : BOOL;
    Error : BOOL;
    ErrorID : UDINT;
END_VAR
VAR
    ax : FB_MotionAxis;
    exPrev : BOOL;
    exEdge : BOOL;
    posAct : DINT;
    np : DINT;
    p : DINT;
END_VAR
    ax.AXIS := Axis;
    exEdge := Execute AND NOT exPrev; exPrev := Execute;
    Busy := FALSE; Done := FALSE; Error := FALSE; ErrorID := 0;
    IF exEdge THEN
        p := LREAL_TO_DINT(Position);
        IF Relative THEN
            np := p;
        ELSE
            ax.OP := 4; ax.INDEX := 16#6064; ax();
            posAct := ax.VALUE;
            np := p - posAct;
        END_IF;
        ax.OP := 5; ax.INDEX := 16#2002; ax.VALUE := np; ax();
        IF ax.STATUS = 0 THEN
            Done := TRUE;
        ELSE
            Error := TRUE; ErrorID := ax.ERRID;
        END_IF;
    END_IF;
END_FUNCTION_BLOCK

// FB_CoEAX8000DeletePositionOffset — clear AX8000 offset (0x2002).
FUNCTION_BLOCK FB_CoEAX8000DeletePositionOffset
VAR_INPUT
    Execute : BOOL;
    Position : LREAL;
    Relative : BOOL;
    Feedback : UDINT;
    Memory : UDINT;
    NetId : STRING[15];
    Axis : UDINT;
END_VAR
VAR_OUTPUT
    Busy : BOOL;
    Done : BOOL;
    Error : BOOL;
    ErrorID : UDINT;
END_VAR
VAR
    ax : FB_MotionAxis;
    exPrev : BOOL;
    exEdge : BOOL;
END_VAR
    ax.AXIS := Axis;
    exEdge := Execute AND NOT exPrev; exPrev := Execute;
    Busy := FALSE; Done := FALSE; Error := FALSE; ErrorID := 0;
    IF exEdge THEN
        ax.OP := 5; ax.INDEX := 16#2002; ax.VALUE := 0; ax();
        IF ax.STATUS = 0 THEN
            Done := TRUE;
        ELSE
            Error := TRUE; ErrorID := ax.ERRID;
        END_IF;
    END_IF;
END_FUNCTION_BLOCK

// FB_CoEAX8000ParkAxis — AX8000 park via CoE object 0x2004.
FUNCTION_BLOCK FB_CoEAX8000ParkAxis
VAR_INPUT
    Execute : BOOL;
    Mode : UDINT;
    NetId : STRING[15];
    Axis : UDINT;
END_VAR
VAR_OUTPUT
    Busy : BOOL;
    Done : BOOL;
    Error : BOOL;
    ErrorID : UDINT;
END_VAR
VAR
    ax : FB_MotionAxis;
    exPrev : BOOL;
    exEdge : BOOL;
END_VAR
    ax.AXIS := Axis;
    exEdge := Execute AND NOT exPrev; exPrev := Execute;
    Busy := FALSE; Done := FALSE; Error := FALSE; ErrorID := 0;
    IF exEdge THEN
        ax.OP := 5; ax.INDEX := 16#2004;
        IF Mode <> 0 THEN ax.VALUE := 1; ELSE ax.VALUE := 0; END_IF;
        ax();
        IF ax.STATUS = 0 THEN
            Done := TRUE;
        ELSE
            Error := TRUE; ErrorID := ax.ERRID;
        END_IF;
    END_IF;
END_FUNCTION_BLOCK

// ================================================================== //
// §4.6 EL72xx CoE — brake/offset over the same OD objects.
// ================================================================== //

// FB_CoEEL72xxBrakeControl — EL72xx brake (OD 0x2003).
FUNCTION_BLOCK FB_CoEEL72xxBrakeControl
VAR_INPUT
    Execute : BOOL;
    Mode : UDINT;
    Axis : UDINT;
END_VAR
VAR_OUTPUT
    Busy : BOOL;
    Done : BOOL;
    Error : BOOL;
    ErrorID : UDINT;
END_VAR
VAR
    ax : FB_MotionAxis;
    exPrev : BOOL;
    exEdge : BOOL;
END_VAR
    ax.AXIS := Axis;
    exEdge := Execute AND NOT exPrev; exPrev := Execute;
    Busy := FALSE; Done := FALSE; Error := FALSE; ErrorID := 0;
    IF exEdge THEN
        ax.OP := 5; ax.INDEX := 16#2003;
        ax.VALUE := UDINT_TO_DINT(Mode); ax();
        IF ax.STATUS = 0 THEN
            Done := TRUE;
        ELSE
            Error := TRUE; ErrorID := ax.ERRID;
        END_IF;
    END_IF;
END_FUNCTION_BLOCK

// FB_CoEEL72xxSetPositionOffset — EL72xx offset (0x2002).
FUNCTION_BLOCK FB_CoEEL72xxSetPositionOffset
VAR_INPUT
    Execute : BOOL;
    Position : LREAL;
    Relative : BOOL;
    Feedback : UDINT;
    Memory : UDINT;
    Axis : UDINT;
END_VAR
VAR_OUTPUT
    Busy : BOOL;
    Done : BOOL;
    Error : BOOL;
    ErrorID : UDINT;
END_VAR
VAR
    ax : FB_MotionAxis;
    exPrev : BOOL;
    exEdge : BOOL;
    posAct : DINT;
    np : DINT;
    p : DINT;
END_VAR
    ax.AXIS := Axis;
    exEdge := Execute AND NOT exPrev; exPrev := Execute;
    Busy := FALSE; Done := FALSE; Error := FALSE; ErrorID := 0;
    IF exEdge THEN
        p := LREAL_TO_DINT(Position);
        IF Relative THEN
            np := p;
        ELSE
            ax.OP := 4; ax.INDEX := 16#6064; ax();
            posAct := ax.VALUE;
            np := p - posAct;
        END_IF;
        ax.OP := 5; ax.INDEX := 16#2002; ax.VALUE := np; ax();
        IF ax.STATUS = 0 THEN
            Done := TRUE;
        ELSE
            Error := TRUE; ErrorID := ax.ERRID;
        END_IF;
    END_IF;
END_FUNCTION_BLOCK

// FB_CoEEL72xxDeletePositionOffset — clear EL72xx offset (0x2002).
FUNCTION_BLOCK FB_CoEEL72xxDeletePositionOffset
VAR_INPUT
    Execute : BOOL;
    Position : LREAL;
    Relative : BOOL;
    Feedback : UDINT;
    Memory : UDINT;
    Axis : UDINT;
END_VAR
VAR_OUTPUT
    Busy : BOOL;
    Done : BOOL;
    Error : BOOL;
    ErrorID : UDINT;
END_VAR
VAR
    ax : FB_MotionAxis;
    exPrev : BOOL;
    exEdge : BOOL;
END_VAR
    ax.AXIS := Axis;
    exEdge := Execute AND NOT exPrev; exPrev := Execute;
    Busy := FALSE; Done := FALSE; Error := FALSE; ErrorID := 0;
    IF exEdge THEN
        ax.OP := 5; ax.INDEX := 16#2002; ax.VALUE := 0; ax();
        IF ax.STATUS = 0 THEN
            Done := TRUE;
        ELSE
            Error := TRUE; ErrorID := ax.ERRID;
        END_IF;
    END_IF;
END_FUNCTION_BLOCK

// ================================================================== //
// §5 Motion blocks
// ================================================================== //

// MC_GearInVelo — velocity-ratio gear coupling (same model as
// MC_GearIn in tc2_mc2.st): slave runs ProfileVelocity at
// master VelocityActualValue * RatioNumerator / RatioDenominator.
// StartSync reports once the slave is tracking (InGear).
FUNCTION_BLOCK MC_GearInVelo
VAR_INPUT
    Execute : BOOL;
    RatioNumerator : DINT;
    RatioDenominator : DINT;
    Acceleration : DINT;
    Deceleration : DINT;
    Master : UDINT;
    Slave : UDINT;
END_VAR
VAR_OUTPUT
    StartSync : BOOL;
    InGear : BOOL;
    Busy : BOOL;
    Error : BOOL;
    ErrorID : UDINT;
END_VAR
VAR
    axM : FB_MotionAxis;
    axS : FB_MotionAxis;
    exPrev : BOOL;
    exEdge : BOOL;
    mvel : DINT;
END_VAR
    axM.AXIS := Master;
    axS.AXIS := Slave;
    axM.OP := 3; axM();
    exEdge := Execute AND NOT exPrev; exPrev := Execute;
    InGear := FALSE;
    Error := FALSE; ErrorID := 0;
    IF exEdge THEN
        IF RatioDenominator = 0 THEN
            Error := TRUE; ErrorID := 1;
        ELSE
            axS.OP := 5; axS.INDEX := 16#6040; axS.VALUE := 16#000F; axS();
            axS.OP := 5; axS.INDEX := 16#6060; axS.VALUE := 3; axS();
        END_IF;
    END_IF;
    IF Execute AND RatioDenominator <> 0 THEN
        axM.OP := 4; axM.INDEX := 16#606C; axM();
        mvel := axM.VALUE;
        axS.OP := 5; axS.INDEX := 16#60FF;
        axS.VALUE := mvel * RatioNumerator / RatioDenominator; axS();
        axS.OP := 6; axS();
        IF axS.STATUS < 0 THEN
            Error := TRUE; ErrorID := axS.ERRID;
        ELSE
            InGear := TRUE;
        END_IF;
    END_IF;
    StartSync := InGear;
    Busy := Execute AND (RatioDenominator <> 0);
END_FUNCTION_BLOCK

// MC_GearInPos — position-ratio master/slave coupling: the slave
// tracks master PositionActualValue * RatioNumerator /
// RatioDenominator through CSP setpoints (0x607A).  Engage edge
// enables the slave and selects CSP mode; release leaves the last
// setpoint (stop via MC_Halt/MC_Stop).  Approximates TwinCAT's
// sync-point gearing with a continuous position ratio — no
// acceleration-profile or sync-window handling.
FUNCTION_BLOCK MC_GearInPos
VAR_INPUT
    Execute : BOOL;
    RatioNumerator : DINT;
    RatioDenominator : DINT;
    Acceleration : DINT;
    Deceleration : DINT;
    Master : UDINT;
    Slave : UDINT;
END_VAR
VAR_OUTPUT
    StartSync : BOOL;
    InGear : BOOL;
    Busy : BOOL;
    CommandAborted : BOOL;
    Error : BOOL;
    ErrorID : UDINT;
END_VAR
VAR
    axM : FB_MotionAxis;
    axS : FB_MotionAxis;
    exPrev : BOOL;
    exEdge : BOOL;
    mpos : DINT;
END_VAR
    axM.AXIS := Master;
    axS.AXIS := Slave;
    axM.OP := 3; axM();
    exEdge := Execute AND NOT exPrev; exPrev := Execute;
    InGear := FALSE;
    CommandAborted := FALSE; Error := FALSE; ErrorID := 0;
    IF exEdge THEN
        IF RatioDenominator = 0 THEN
            Error := TRUE; ErrorID := 1;
        ELSE
            axS.OP := 5; axS.INDEX := 16#6040; axS.VALUE := 16#000F; axS();
            axS.OP := 5; axS.INDEX := 16#6060; axS.VALUE := 8; axS();
        END_IF;
    END_IF;
    IF Execute AND RatioDenominator <> 0 THEN
        axM.OP := 4; axM.INDEX := 16#6064; axM();
        mpos := axM.VALUE;
        axS.OP := 5; axS.INDEX := 16#607A;
        axS.VALUE := mpos * RatioNumerator / RatioDenominator; axS();
        axS.OP := 6; axS();
        IF axS.STATUS < 0 THEN
            Error := TRUE; ErrorID := axS.ERRID;
        ELSE
            InGear := TRUE;
        END_IF;
    END_IF;
    StartSync := InGear;
    Busy := Execute AND (RatioDenominator <> 0);
END_FUNCTION_BLOCK

// MC_ReadFlyingSawCharacteristics — read the flying-saw
// characteristic values (OD 0x2006..0x2009 -> Value0..Value3).
// CamTableCharac is flattened to four DINT outputs.
FUNCTION_BLOCK MC_ReadFlyingSawCharacteristics
VAR_INPUT
    Execute : BOOL;
    Slave : UDINT;
END_VAR
VAR_OUTPUT
    Value0 : DINT;
    Value1 : DINT;
    Value2 : DINT;
    Value3 : DINT;
    Busy : BOOL;
    Done : BOOL;
    Error : BOOL;
    ErrorID : UDINT;
END_VAR
VAR
    ax : FB_MotionAxis;
    exPrev : BOOL;
    exEdge : BOOL;
    i : DINT;
END_VAR
    ax.AXIS := Slave;
    exEdge := Execute AND NOT exPrev; exPrev := Execute;
    Busy := FALSE; Done := FALSE; Error := FALSE; ErrorID := 0;
    IF exEdge THEN
        FOR i := 0 TO 3 DO
            ax.OP := 4;
            ax.INDEX := 16#2006 + i;
            ax();
            IF ax.STATUS <> 0 THEN
                Error := TRUE; ErrorID := ax.ERRID;
            ELSIF i = 0 THEN Value0 := ax.VALUE;
            ELSIF i = 1 THEN Value1 := ax.VALUE;
            ELSIF i = 2 THEN Value2 := ax.VALUE;
            ELSE Value3 := ax.VALUE;
            END_IF;
        END_FOR;
        IF NOT Error THEN Done := TRUE; END_IF;
    END_IF;
END_FUNCTION_BLOCK

// ---- version --------------------------------------------------------

// F_GetVersionTcMc2Drive — library version placeholder.
FUNCTION F_GetVersionTcMc2Drive : UDINT
F_GetVersionTcMc2Drive := 16#0100;
END_FUNCTION

(* ---- tc2_mc2_xfc.st ---- *)
// Tc2_MC2_XFC + Tc2_NciXFC + Tc3_MC2_AdvancedHoming_XFC (subset)
// XFC cyclic setpoint evaluation over FB_MotionAxis.
//
// Time base: each FB owns a TON clock (IN held TRUE) whose ET is the
// nanosecond scan clock; DC time is flattened to the low 32 bits of
// that clock (T_DCTIME32 semantics, wraps at ~4.29 s).  Axis
// kinematics use the OP6 snapshot (POS_ACTUAL/VEL_ACTUAL, user
// units, velocity in user units per second) with linear
// extrapolation — the real XFC kernel evaluates the full motion
// profile, so trapezoid/segment extrapolation is a documented gap.
// AXIS_REF is the UDINT handle; OUTPUT_REF/CAMSWITCH_REF/TRACK_REF
// and the EL terminal structs are flattened to BOOL/LREAL members.

// Shared clock helper: TON ET is ns; expose low32 as UDINT.
FUNCTION_BLOCK XFC_Clock
VAR_OUTPUT
    DcTime : UDINT;   // low 32 bits of the ns scan clock
    NowNs  : LINT;    // full ns (may exceed 32 bits on long runs)
END_VAR
VAR
    clk : TON;
END_VAR
    clk(IN := TRUE, PT := T#1000000h);
    DcTime := TIME_TO_UDINT(clk.ET);
    NowNs := TIME_TO_LINT(clk.ET);
END_FUNCTION_BLOCK

// XFC_PositionAtTime — extrapolated axis position at DcTime.
FUNCTION_BLOCK XFC_PositionAtTime
VAR_INPUT
    DcTime : UDINT;
    Axis   : UDINT;
END_VAR
VAR_OUTPUT
    Position : LREAL;
    Error    : BOOL;
    ErrorID  : UDINT;
END_VAR
VAR
    clk : XFC_Clock;
    ax  : FB_MotionAxis;
    dt  : DINT;
    pos : DINT;
    vel : DINT;
END_VAR
    clk();
    ax.AXIS := Axis;
    ax.OP := 6; ax();
    Error := FALSE; ErrorID := 0;
    IF ax.STATUS < 0 THEN
        Error := TRUE; ErrorID := ax.ERRID;
    ELSE
        pos := ax.POS_ACTUAL;
        vel := ax.VEL_ACTUAL;
        // 32-bit modular delta, interpreted signed (ns)
        dt := UDINT_TO_DINT(DcTime - clk.DcTime);
        Position := DINT_TO_LREAL(pos)
                  + DINT_TO_LREAL(vel) * DINT_TO_LREAL(dt) / 1000000000.0;
    END_IF;
END_FUNCTION_BLOCK

// XFC_TimeOfPosition — DC time at which the axis reaches Position.
FUNCTION_BLOCK XFC_TimeOfPosition
VAR_INPUT
    Position : LREAL;
    Axis     : UDINT;
END_VAR
VAR_OUTPUT
    DcTime  : UDINT;
    Error   : BOOL;
    ErrorID : UDINT;
END_VAR
VAR
    clk : XFC_Clock;
    ax  : FB_MotionAxis;
    pos : DINT;
    vel : DINT;
    dtNs : LREAL;
END_VAR
    clk();
    ax.AXIS := Axis;
    ax.OP := 6; ax();
    Error := FALSE; ErrorID := 0; DcTime := clk.DcTime;
    IF ax.STATUS < 0 THEN
        Error := TRUE; ErrorID := ax.ERRID;
    ELSE
        pos := ax.POS_ACTUAL;
        vel := ax.VEL_ACTUAL;
        IF vel <> 0 THEN
            dtNs := (Position - DINT_TO_LREAL(pos))
                    / DINT_TO_LREAL(vel) * 1000000000.0;
            DcTime := clk.DcTime + LREAL_TO_UDINT(dtNs);
        END_IF;
    END_IF;
END_FUNCTION_BLOCK

// XFC_TimeToPosition — signed ns until the axis reaches Position
// (negative when the position is in the past).
FUNCTION_BLOCK XFC_TimeToPosition
VAR_INPUT
    Position : LREAL;
    Axis     : UDINT;
END_VAR
VAR_OUTPUT
    Duration : DINT;
    Error    : BOOL;
    ErrorID  : UDINT;
END_VAR
VAR
    clk : XFC_Clock;
    ax  : FB_MotionAxis;
    pos : DINT;
    vel : DINT;
END_VAR
    clk();
    ax.AXIS := Axis;
    ax.OP := 6; ax();
    Error := FALSE; ErrorID := 0; Duration := 0;
    IF ax.STATUS < 0 THEN
        Error := TRUE; ErrorID := ax.ERRID;
    ELSE
        pos := ax.POS_ACTUAL;
        vel := ax.VEL_ACTUAL;
        IF vel <> 0 THEN
            Duration := LREAL_TO_DINT((Position - DINT_TO_LREAL(pos))
                             / DINT_TO_LREAL(vel) * 1000000000.0);
        END_IF;
    END_IF;
END_FUNCTION_BLOCK

// XFC_TimeToModuloPosition — time to the nearest modulo position in
// the direction of travel.  ModuloFactor is the position wrap
// (0 disables wrapping).
FUNCTION_BLOCK XFC_TimeToModuloPosition
VAR_INPUT
    Position      : LREAL;
    ModuloFactor  : LREAL;
    Axis          : UDINT;
END_VAR
VAR_OUTPUT
    Duration : DINT;
    Error    : BOOL;
    ErrorID  : UDINT;
END_VAR
VAR
    clk : XFC_Clock;
    ax  : FB_MotionAxis;
    pos : DINT;
    vel : DINT;
    p   : LREAL;
END_VAR
    clk();
    ax.AXIS := Axis;
    ax.OP := 6; ax();
    Error := FALSE; ErrorID := 0; Duration := 0;
    IF ax.STATUS < 0 THEN
        Error := TRUE; ErrorID := ax.ERRID;
    ELSE
        pos := ax.POS_ACTUAL;
        vel := ax.VEL_ACTUAL;
        p := Position;
        IF ModuloFactor > 0.0 THEN
            // wrap target into the revolution around pos
            WHILE p < DINT_TO_LREAL(pos) - ModuloFactor / 2.0 DO
                p := p + ModuloFactor;
            END_WHILE;
            WHILE p > DINT_TO_LREAL(pos) + ModuloFactor / 2.0 DO
                p := p - ModuloFactor;
            END_WHILE;
        END_IF;
        IF vel <> 0 THEN
            Duration := LREAL_TO_DINT((p - DINT_TO_LREAL(pos))
                             / DINT_TO_LREAL(vel) * 1000000000.0);
        END_IF;
    END_IF;
END_FUNCTION_BLOCK

// XFC_GetCurDcTaskTime — current DC task time (low32 of the ns
// clock; the FUNCTION form is flattened to an FB).
FUNCTION_BLOCK XFC_GetCurDcTaskTime
VAR_OUTPUT
    DcTime : UDINT;
END_VAR
VAR
    clk : XFC_Clock;
END_VAR
    clk();
    DcTime := clk.DcTime;
END_FUNCTION_BLOCK

// XFC_ExtendDcTime — extend a 32-bit DC time against a reference.
// The sim clock domain is 32-bit, so the FB reports the signed
// nanosecond offset of DcTime32 relative to RefDcTime (the 64-bit
// T_DCTIME result cannot be represented).
FUNCTION_BLOCK XFC_ExtendDcTime
VAR_INPUT
    DcTime32  : UDINT;
    RefDcTime : UDINT;
END_VAR
VAR_OUTPUT
    DeltaNs : DINT;
    DcTime  : UDINT;
END_VAR
    DeltaNs := UDINT_TO_DINT(DcTime32 - RefDcTime);
    DcTime := DcTime32;
END_FUNCTION_BLOCK

// XFC_PositionCam — digital output on inside [FirstOn,LastOn].
// OUTPUT_REF flattened to a BOOL output; Modulo wraps positions by
// ModuloFactor (0 = absolute).
FUNCTION_BLOCK XFC_PositionCam
VAR_INPUT
    FirstOnPosition : LREAL;
    LastOnPosition  : LREAL;
    Modulo          : BOOL;
    ModuloFactor    : LREAL;
    Axis            : UDINT;
END_VAR
VAR_OUTPUT
    Output  : BOOL;
    Error   : BOOL;
    ErrorID : UDINT;
END_VAR
VAR
    ax  : FB_MotionAxis;
    pos : LREAL;
    p   : LREAL;
END_VAR
    ax.AXIS := Axis;
    ax.OP := 6; ax();
    Error := FALSE; ErrorID := 0; Output := FALSE;
    IF ax.STATUS < 0 THEN
        Error := TRUE; ErrorID := ax.ERRID;
    ELSE
        pos := DINT_TO_LREAL(ax.POS_ACTUAL);
        p := pos;
        IF Modulo AND ModuloFactor > 0.0 THEN
            p := pos - DINT_TO_LREAL(LREAL_TO_DINT(pos / ModuloFactor)) * ModuloFactor;
        END_IF;
        IF p >= FirstOnPosition AND p <= LastOnPosition THEN
            Output := TRUE;
        END_IF;
    END_IF;
END_FUNCTION_BLOCK

// XFC_TimeCam — output ON from FirstOnPosition for Duration
// seconds (position-triggered, time-limited).
FUNCTION_BLOCK XFC_TimeCam
VAR_INPUT
    FirstOnPosition : LREAL;
    Duration        : LREAL;
    Modulo          : BOOL;
    ModuloFactor    : LREAL;
    Axis            : UDINT;
END_VAR
VAR_OUTPUT
    Output  : BOOL;
    Error   : BOOL;
    ErrorID : UDINT;
END_VAR
VAR
    clk   : XFC_Clock;
    ax    : FB_MotionAxis;
    pos   : LREAL;
    p     : LREAL;
    armed : BOOL;
    onAt  : LINT;
END_VAR
    clk();
    ax.AXIS := Axis;
    ax.OP := 6; ax();
    Error := FALSE; ErrorID := 0; Output := FALSE;
    IF ax.STATUS < 0 THEN
        Error := TRUE; ErrorID := ax.ERRID;
    ELSE
        pos := DINT_TO_LREAL(ax.POS_ACTUAL);
        p := pos;
        IF Modulo AND ModuloFactor > 0.0 THEN
            p := pos - DINT_TO_LREAL(LREAL_TO_DINT(pos / ModuloFactor)) * ModuloFactor;
        END_IF;
        // one shot per crossing: re-arms only when position drops
        // back below FirstOnPosition
        IF p < FirstOnPosition THEN
            armed := FALSE;
        ELSIF p >= FirstOnPosition AND NOT armed THEN
            armed := TRUE;
            onAt := clk.NowNs;
        END_IF;
        IF armed AND (LINT_TO_LREAL(clk.NowNs - onAt) / 1000000000.0) < Duration THEN
            Output := TRUE;
        END_IF;
    END_IF;
END_FUNCTION_BLOCK

// XFC_BreakCam — brake cam: Output follows BreakRelease while the
// axis is valid (the position-dependent release curve of the real
// block is not modeled).
FUNCTION_BLOCK XFC_BreakCam
VAR_INPUT
    BreakRelease : BOOL;
    Axis         : UDINT;
END_VAR
VAR_OUTPUT
    Output  : BOOL;
    Error   : BOOL;
    ErrorID : UDINT;
END_VAR
VAR
    ax : FB_MotionAxis;
END_VAR
    ax.AXIS := Axis;
    ax.OP := 6; ax();
    Error := FALSE; ErrorID := 0;
    IF ax.STATUS < 0 THEN
        Error := TRUE; ErrorID := ax.ERRID;
    ELSE
        Output := BreakRelease;
    END_IF;
END_FUNCTION_BLOCK

// MC_DigitalCamSwitch — single-cam digital switch (CAMSWITCH_REF/
// OUTPUT_REF/TRACK_REF flattened to FirstOn/LastOn/Modulo + BOOL).
// MC_DigitalCamSwitch_MultiEdge shares this implementation.
FUNCTION_BLOCK MC_DigitalCamSwitch
VAR_INPUT
    Enable          : BOOL;
    FirstOnPosition : LREAL;
    LastOnPosition  : LREAL;
    Modulo          : BOOL;
    ModuloFactor    : LREAL;
    Axis            : UDINT;
END_VAR
VAR_OUTPUT
    InOperation : BOOL;
    Output      : BOOL;
    Error       : BOOL;
    ErrorID     : UDINT;
END_VAR
VAR
    cam : XFC_PositionCam;
END_VAR
    InOperation := Enable;
    cam(FirstOnPosition := FirstOnPosition,
        LastOnPosition  := LastOnPosition,
        Modulo          := Modulo,
        ModuloFactor    := ModuloFactor,
        Axis            := Axis);
    Output := Enable AND cam.Output;
    Error := cam.Error;
    ErrorID := cam.ErrorID;
END_FUNCTION_BLOCK

// MC_DigitalCamSwitch_MultiEdge — same flattened single-cam model;
// the multi-edge/EL5131 track variant is not modeled.
FUNCTION_BLOCK MC_DigitalCamSwitch_MultiEdge
VAR_INPUT
    Enable          : BOOL;
    FirstOnPosition : LREAL;
    LastOnPosition  : LREAL;
    Modulo          : BOOL;
    ModuloFactor    : LREAL;
    Axis            : UDINT;
END_VAR
VAR_OUTPUT
    InOperation : BOOL;
    Output      : BOOL;
    Error       : BOOL;
    ErrorID     : UDINT;
END_VAR
VAR
    cam : XFC_PositionCam;
END_VAR
    InOperation := Enable;
    cam(FirstOnPosition := FirstOnPosition,
        LastOnPosition  := LastOnPosition,
        Modulo          := Modulo,
        ModuloFactor    := ModuloFactor,
        Axis            := Axis);
    Output := Enable AND cam.Output;
    Error := cam.Error;
    ErrorID := cam.ErrorID;
END_FUNCTION_BLOCK

// XFC_TouchProbe — record PositionActualValue on the TriggerInput
// rising edge while Execute is active (XFC_TRIGGER_REF flattened
// to BOOL).
FUNCTION_BLOCK XFC_TouchProbe
VAR_INPUT
    Execute       : BOOL;
    TriggerInput  : BOOL;
    Axis          : UDINT;
END_VAR
VAR_OUTPUT
    RecordedPosition : LREAL;
    Done             : BOOL;
    Busy             : BOOL;
    Error            : BOOL;
    ErrorID          : UDINT;
END_VAR
VAR
    ax        : FB_MotionAxis;
    exPrev    : BOOL;
    exEdge    : BOOL;
    trgPrev   : BOOL;
    armed     : BOOL;
END_VAR
    ax.AXIS := Axis;
    exEdge := Execute AND NOT exPrev; exPrev := Execute;
    Busy := FALSE; Done := FALSE; Error := FALSE; ErrorID := 0;
    IF exEdge THEN
        armed := TRUE;
    END_IF;
    IF NOT Execute THEN armed := FALSE; END_IF;
    IF armed AND TriggerInput AND NOT trgPrev THEN
        ax.OP := 6; ax();
        IF ax.STATUS < 0 THEN
            Error := TRUE; ErrorID := ax.ERRID;
        ELSE
            RecordedPosition := DINT_TO_LREAL(ax.POS_ACTUAL);
            Done := TRUE;
            armed := FALSE;
        END_IF;
    END_IF;
    Busy := armed;
    trgPrev := TriggerInput;
END_FUNCTION_BLOCK

// ---- version --------------------------------------------------------

// F_GetVersionTcXfc — library version placeholder.
FUNCTION F_GetVersionTcXfc : UDINT
F_GetVersionTcXfc := 16#0100;
END_FUNCTION

(* ---- tc2_modbusrtu.st ---- *)
// Tc2_ModbusRTU Modbus RTU master FBs (TwinCAT 3 PLC Library
// Tc2_ModbusRTU, manual TF6255). Beckhoff-shaped wrappers over the
// builtin FB_ModbusRtu, which drives the host "tplc-modbus" service
// RTU transport (serial device opened per transaction, RTU framing
// unit|func|data|crc16, CRC-validated responses, nonblocking).
// TwinCAT exposes each Modbus function as an action on the
// ModbusRtuMasterV2_* FBs; here each action is a standalone FB with
// the same parameters. Differences from TwinCAT, documented in
// docs/plc/compat/README.md:
//   - POINTER TO BYTE payloads are ARRAY[0..255] OF BYTE buffers
//     (bounded; cbLength/cbSrcLength/cbDestLength still apply).
//   - serial line settings are explicit inputs (sDevice, nBaud,
//     nParity, nDataBits, nStopBits) instead of TwinCAT System
//     Manager COM-port bindings.
//   - nErrId carries tplc-modbus transport codes, or the Modbus
//     exception code when the slave returns an exception response.
//   - ModbusRtuSlave_* and the *_Generic ComBuffer variants are not
//     provided; KL6x*B bus-terminal variants need EtherCAT terminal
//     integration.
// Sources: docs/plc/plan/21-twincat-libraries.md §7 (TF6255).

FUNCTION_BLOCK FB_MBRtuReadCoils
VAR_INPUT
    sDevice : STRING[63];
    nBaud : UDINT := 9600;
    nParity : UDINT := 0;
    nDataBits : UDINT := 8;
    nStopBits : UDINT := 1;
    nUnitID : BYTE := 1;
    nQuantity : WORD;
    nMBAddr : WORD;
    cbLength : UDINT;
    bExecute : BOOL;
    tTimeout : TIME;
END_VAR
VAR_OUTPUT
    bBusy : BOOL;
    bDone : BOOL;
    bError : BOOL;
    nErrId : UDINT;
    cbRead : UDINT;
    pData : ARRAY[0..255] OF BYTE;
END_VAR
VAR
    mb : FB_ModbusRtu;
    i : UDINT;
END_VAR
    mb.FUNC := 1;
    mb.DEV := sDevice;
    mb.BAUD := nBaud;
    mb.PARITY := nParity;
    mb.DBITS := nDataBits;
    mb.SBITS := nStopBits;
    mb.UNIT := nUnitID;
    mb.TIMEOUT := tTimeout;
    mb.DATA[0] := UINT_TO_BYTE(nMBAddr / 256);
    mb.DATA[1] := UINT_TO_BYTE(nMBAddr MOD 256);
    mb.DATA[2] := UINT_TO_BYTE(nQuantity / 256);
    mb.DATA[3] := UINT_TO_BYTE(nQuantity MOD 256);
    mb.RLEN := 4;
    mb.EXEC := bExecute;
    mb();
    bBusy := mb.BUSY;
    bDone := mb.DONE;
    IF mb.DONE THEN
        i := 0;
        WHILE i < mb.DLEN AND i < 256 DO
            pData[i] := mb.DATA[i];
            i := i + 1;
        END_WHILE;
        cbRead := mb.DLEN;
    END_IF;
    nErrId := mb.ERRID;
    IF mb.RESULT = 1 THEN
        nErrId := 16#8000 + mb.EXC;
    END_IF;
    bError := (mb.ERRID <> 0) OR (mb.RESULT = 1);
END_FUNCTION_BLOCK

FUNCTION_BLOCK FB_MBRtuReadInputs
VAR_INPUT
    sDevice : STRING[63];
    nBaud : UDINT := 9600;
    nParity : UDINT := 0;
    nDataBits : UDINT := 8;
    nStopBits : UDINT := 1;
    nUnitID : BYTE := 1;
    nQuantity : WORD;
    nMBAddr : WORD;
    cbLength : UDINT;
    bExecute : BOOL;
    tTimeout : TIME;
END_VAR
VAR_OUTPUT
    bBusy : BOOL;
    bDone : BOOL;
    bError : BOOL;
    nErrId : UDINT;
    cbRead : UDINT;
    pData : ARRAY[0..255] OF BYTE;
END_VAR
VAR
    mb : FB_ModbusRtu;
    i : UDINT;
END_VAR
    mb.FUNC := 2;
    mb.DEV := sDevice;
    mb.BAUD := nBaud;
    mb.PARITY := nParity;
    mb.DBITS := nDataBits;
    mb.SBITS := nStopBits;
    mb.UNIT := nUnitID;
    mb.TIMEOUT := tTimeout;
    mb.DATA[0] := UINT_TO_BYTE(nMBAddr / 256);
    mb.DATA[1] := UINT_TO_BYTE(nMBAddr MOD 256);
    mb.DATA[2] := UINT_TO_BYTE(nQuantity / 256);
    mb.DATA[3] := UINT_TO_BYTE(nQuantity MOD 256);
    mb.RLEN := 4;
    mb.EXEC := bExecute;
    mb();
    bBusy := mb.BUSY;
    bDone := mb.DONE;
    IF mb.DONE THEN
        i := 0;
        WHILE i < mb.DLEN AND i < 256 DO
            pData[i] := mb.DATA[i];
            i := i + 1;
        END_WHILE;
        cbRead := mb.DLEN;
    END_IF;
    nErrId := mb.ERRID;
    IF mb.RESULT = 1 THEN
        nErrId := 16#8000 + mb.EXC;
    END_IF;
    bError := (mb.ERRID <> 0) OR (mb.RESULT = 1);
END_FUNCTION_BLOCK

FUNCTION_BLOCK FB_MBRtuReadRegs
VAR_INPUT
    sDevice : STRING[63];
    nBaud : UDINT := 9600;
    nParity : UDINT := 0;
    nDataBits : UDINT := 8;
    nStopBits : UDINT := 1;
    nUnitID : BYTE := 1;
    nQuantity : WORD;
    nMBAddr : WORD;
    cbLength : UDINT;
    bExecute : BOOL;
    tTimeout : TIME;
END_VAR
VAR_OUTPUT
    bBusy : BOOL;
    bDone : BOOL;
    bError : BOOL;
    nErrId : UDINT;
    cbRead : UDINT;
    pData : ARRAY[0..255] OF BYTE;
END_VAR
VAR
    mb : FB_ModbusRtu;
    i : UDINT;
END_VAR
    mb.FUNC := 3;
    mb.DEV := sDevice;
    mb.BAUD := nBaud;
    mb.PARITY := nParity;
    mb.DBITS := nDataBits;
    mb.SBITS := nStopBits;
    mb.UNIT := nUnitID;
    mb.TIMEOUT := tTimeout;
    mb.DATA[0] := UINT_TO_BYTE(nMBAddr / 256);
    mb.DATA[1] := UINT_TO_BYTE(nMBAddr MOD 256);
    mb.DATA[2] := UINT_TO_BYTE(nQuantity / 256);
    mb.DATA[3] := UINT_TO_BYTE(nQuantity MOD 256);
    mb.RLEN := 4;
    mb.EXEC := bExecute;
    mb();
    bBusy := mb.BUSY;
    bDone := mb.DONE;
    IF mb.DONE THEN
        i := 0;
        WHILE i < mb.DLEN AND i < 256 DO
            pData[i] := mb.DATA[i];
            i := i + 1;
        END_WHILE;
        cbRead := mb.DLEN;
    END_IF;
    nErrId := mb.ERRID;
    IF mb.RESULT = 1 THEN
        nErrId := 16#8000 + mb.EXC;
    END_IF;
    bError := (mb.ERRID <> 0) OR (mb.RESULT = 1);
END_FUNCTION_BLOCK

FUNCTION_BLOCK FB_MBRtuReadInputRegs
VAR_INPUT
    sDevice : STRING[63];
    nBaud : UDINT := 9600;
    nParity : UDINT := 0;
    nDataBits : UDINT := 8;
    nStopBits : UDINT := 1;
    nUnitID : BYTE := 1;
    nQuantity : WORD;
    nMBAddr : WORD;
    cbLength : UDINT;
    bExecute : BOOL;
    tTimeout : TIME;
END_VAR
VAR_OUTPUT
    bBusy : BOOL;
    bDone : BOOL;
    bError : BOOL;
    nErrId : UDINT;
    cbRead : UDINT;
    pData : ARRAY[0..255] OF BYTE;
END_VAR
VAR
    mb : FB_ModbusRtu;
    i : UDINT;
END_VAR
    mb.FUNC := 4;
    mb.DEV := sDevice;
    mb.BAUD := nBaud;
    mb.PARITY := nParity;
    mb.DBITS := nDataBits;
    mb.SBITS := nStopBits;
    mb.UNIT := nUnitID;
    mb.TIMEOUT := tTimeout;
    mb.DATA[0] := UINT_TO_BYTE(nMBAddr / 256);
    mb.DATA[1] := UINT_TO_BYTE(nMBAddr MOD 256);
    mb.DATA[2] := UINT_TO_BYTE(nQuantity / 256);
    mb.DATA[3] := UINT_TO_BYTE(nQuantity MOD 256);
    mb.RLEN := 4;
    mb.EXEC := bExecute;
    mb();
    bBusy := mb.BUSY;
    bDone := mb.DONE;
    IF mb.DONE THEN
        i := 0;
        WHILE i < mb.DLEN AND i < 256 DO
            pData[i] := mb.DATA[i];
            i := i + 1;
        END_WHILE;
        cbRead := mb.DLEN;
    END_IF;
    nErrId := mb.ERRID;
    IF mb.RESULT = 1 THEN
        nErrId := 16#8000 + mb.EXC;
    END_IF;
    bError := (mb.ERRID <> 0) OR (mb.RESULT = 1);
END_FUNCTION_BLOCK

FUNCTION_BLOCK FB_MBRtuWriteSingleCoil
VAR_INPUT
    sDevice : STRING[63];
    nBaud : UDINT := 9600;
    nParity : UDINT := 0;
    nDataBits : UDINT := 8;
    nStopBits : UDINT := 1;
    nUnitID : BYTE := 1;
    nMBAddr : WORD;
    nValue : WORD;
    bExecute : BOOL;
    tTimeout : TIME;
END_VAR
VAR_OUTPUT
    bBusy : BOOL;
    bDone : BOOL;
    bError : BOOL;
    nErrId : UDINT;
    cbRead : UDINT;
END_VAR
VAR
    mb : FB_ModbusRtu;
END_VAR
    mb.FUNC := 5;
    mb.DEV := sDevice;
    mb.BAUD := nBaud;
    mb.PARITY := nParity;
    mb.DBITS := nDataBits;
    mb.SBITS := nStopBits;
    mb.UNIT := nUnitID;
    mb.TIMEOUT := tTimeout;
    mb.DATA[0] := UINT_TO_BYTE(nMBAddr / 256);
    mb.DATA[1] := UINT_TO_BYTE(nMBAddr MOD 256);
    mb.DATA[2] := UINT_TO_BYTE(nValue / 256);
    mb.DATA[3] := UINT_TO_BYTE(nValue MOD 256);
    mb.RLEN := 4;
    mb.EXEC := bExecute;
    mb();
    bBusy := mb.BUSY;
    bDone := mb.DONE;
    cbRead := 0;
    nErrId := mb.ERRID;
    IF mb.RESULT = 1 THEN
        nErrId := 16#8000 + mb.EXC;
    END_IF;
    bError := (mb.ERRID <> 0) OR (mb.RESULT = 1);
END_FUNCTION_BLOCK

FUNCTION_BLOCK FB_MBRtuWriteSingleReg
VAR_INPUT
    sDevice : STRING[63];
    nBaud : UDINT := 9600;
    nParity : UDINT := 0;
    nDataBits : UDINT := 8;
    nStopBits : UDINT := 1;
    nUnitID : BYTE := 1;
    nMBAddr : WORD;
    nValue : WORD;
    bExecute : BOOL;
    tTimeout : TIME;
END_VAR
VAR_OUTPUT
    bBusy : BOOL;
    bDone : BOOL;
    bError : BOOL;
    nErrId : UDINT;
    cbRead : UDINT;
END_VAR
VAR
    mb : FB_ModbusRtu;
END_VAR
    mb.FUNC := 6;
    mb.DEV := sDevice;
    mb.BAUD := nBaud;
    mb.PARITY := nParity;
    mb.DBITS := nDataBits;
    mb.SBITS := nStopBits;
    mb.UNIT := nUnitID;
    mb.TIMEOUT := tTimeout;
    mb.DATA[0] := UINT_TO_BYTE(nMBAddr / 256);
    mb.DATA[1] := UINT_TO_BYTE(nMBAddr MOD 256);
    mb.DATA[2] := UINT_TO_BYTE(nValue / 256);
    mb.DATA[3] := UINT_TO_BYTE(nValue MOD 256);
    mb.RLEN := 4;
    mb.EXEC := bExecute;
    mb();
    bBusy := mb.BUSY;
    bDone := mb.DONE;
    cbRead := 0;
    nErrId := mb.ERRID;
    IF mb.RESULT = 1 THEN
        nErrId := 16#8000 + mb.EXC;
    END_IF;
    bError := (mb.ERRID <> 0) OR (mb.RESULT = 1);
END_FUNCTION_BLOCK

FUNCTION_BLOCK FB_MBRtuWriteCoils
VAR_INPUT
    sDevice : STRING[63];
    nBaud : UDINT := 9600;
    nParity : UDINT := 0;
    nDataBits : UDINT := 8;
    nStopBits : UDINT := 1;
    nUnitID : BYTE := 1;
    nQuantity : WORD;
    nMBAddr : WORD;
    cbLength : UDINT;
    pSrcData : ARRAY[0..255] OF BYTE;
    bExecute : BOOL;
    tTimeout : TIME;
END_VAR
VAR_OUTPUT
    bBusy : BOOL;
    bDone : BOOL;
    bError : BOOL;
    nErrId : UDINT;
    cbRead : UDINT;
END_VAR
VAR
    mb : FB_ModbusRtu;
    i : UDINT;
    n : UDINT;
END_VAR
    mb.FUNC := 15;
    mb.DEV := sDevice;
    mb.BAUD := nBaud;
    mb.PARITY := nParity;
    mb.DBITS := nDataBits;
    mb.SBITS := nStopBits;
    mb.UNIT := nUnitID;
    mb.TIMEOUT := tTimeout;
    mb.DATA[0] := UINT_TO_BYTE(nMBAddr / 256);
    mb.DATA[1] := UINT_TO_BYTE(nMBAddr MOD 256);
    mb.DATA[2] := UINT_TO_BYTE(nQuantity / 256);
    mb.DATA[3] := UINT_TO_BYTE(nQuantity MOD 256);
    n := cbLength;
    IF n > 246 THEN
        n := 246;
    END_IF;
    mb.DATA[4] := UDINT_TO_BYTE(n);
    i := 0;
    WHILE i < n DO
        mb.DATA[5 + i] := pSrcData[i];
        i := i + 1;
    END_WHILE;
    mb.RLEN := 5 + n;
    mb.EXEC := bExecute;
    mb();
    bBusy := mb.BUSY;
    bDone := mb.DONE;
    cbRead := 0;
    nErrId := mb.ERRID;
    IF mb.RESULT = 1 THEN
        nErrId := 16#8000 + mb.EXC;
    END_IF;
    bError := (mb.ERRID <> 0) OR (mb.RESULT = 1);
END_FUNCTION_BLOCK

FUNCTION_BLOCK FB_MBRtuWriteRegs
VAR_INPUT
    sDevice : STRING[63];
    nBaud : UDINT := 9600;
    nParity : UDINT := 0;
    nDataBits : UDINT := 8;
    nStopBits : UDINT := 1;
    nUnitID : BYTE := 1;
    nQuantity : WORD;
    nMBAddr : WORD;
    cbLength : UDINT;
    pSrcData : ARRAY[0..255] OF BYTE;
    bExecute : BOOL;
    tTimeout : TIME;
END_VAR
VAR_OUTPUT
    bBusy : BOOL;
    bDone : BOOL;
    bError : BOOL;
    nErrId : UDINT;
    cbRead : UDINT;
END_VAR
VAR
    mb : FB_ModbusRtu;
    i : UDINT;
    n : UDINT;
END_VAR
    mb.FUNC := 16;
    mb.DEV := sDevice;
    mb.BAUD := nBaud;
    mb.PARITY := nParity;
    mb.DBITS := nDataBits;
    mb.SBITS := nStopBits;
    mb.UNIT := nUnitID;
    mb.TIMEOUT := tTimeout;
    mb.DATA[0] := UINT_TO_BYTE(nMBAddr / 256);
    mb.DATA[1] := UINT_TO_BYTE(nMBAddr MOD 256);
    mb.DATA[2] := UINT_TO_BYTE(nQuantity / 256);
    mb.DATA[3] := UINT_TO_BYTE(nQuantity MOD 256);
    n := cbLength;
    IF n > 246 THEN
        n := 246;
    END_IF;
    mb.DATA[4] := UDINT_TO_BYTE(n);
    i := 0;
    WHILE i < n DO
        mb.DATA[5 + i] := pSrcData[i];
        i := i + 1;
    END_WHILE;
    mb.RLEN := 5 + n;
    mb.EXEC := bExecute;
    mb();
    bBusy := mb.BUSY;
    bDone := mb.DONE;
    cbRead := 0;
    nErrId := mb.ERRID;
    IF mb.RESULT = 1 THEN
        nErrId := 16#8000 + mb.EXC;
    END_IF;
    bError := (mb.ERRID <> 0) OR (mb.RESULT = 1);
END_FUNCTION_BLOCK

FUNCTION_BLOCK FB_MBRtuReadWriteRegs
VAR_INPUT
    sDevice : STRING[63];
    nBaud : UDINT := 9600;
    nParity : UDINT := 0;
    nDataBits : UDINT := 8;
    nStopBits : UDINT := 1;
    nUnitID : BYTE := 1;
    nReadQuantity : WORD;
    nMBReadAddr : WORD;
    nWriteQuantity : WORD;
    nMBWriteAddr : WORD;
    cbDestLength : UDINT;
    cbSrcLength : UDINT;
    pSrcData : ARRAY[0..255] OF BYTE;
    bExecute : BOOL;
    tTimeout : TIME;
END_VAR
VAR_OUTPUT
    bBusy : BOOL;
    bDone : BOOL;
    bError : BOOL;
    nErrId : UDINT;
    cbRead : UDINT;
    pDestData : ARRAY[0..255] OF BYTE;
END_VAR
VAR
    mb : FB_ModbusRtu;
    i : UDINT;
    n : UDINT;
END_VAR
    mb.FUNC := 23;
    mb.DEV := sDevice;
    mb.BAUD := nBaud;
    mb.PARITY := nParity;
    mb.DBITS := nDataBits;
    mb.SBITS := nStopBits;
    mb.UNIT := nUnitID;
    mb.TIMEOUT := tTimeout;
    mb.DATA[0] := UINT_TO_BYTE(nMBReadAddr / 256);
    mb.DATA[1] := UINT_TO_BYTE(nMBReadAddr MOD 256);
    mb.DATA[2] := UINT_TO_BYTE(nReadQuantity / 256);
    mb.DATA[3] := UINT_TO_BYTE(nReadQuantity MOD 256);
    mb.DATA[4] := UINT_TO_BYTE(nMBWriteAddr / 256);
    mb.DATA[5] := UINT_TO_BYTE(nMBWriteAddr MOD 256);
    mb.DATA[6] := UINT_TO_BYTE(nWriteQuantity / 256);
    mb.DATA[7] := UINT_TO_BYTE(nWriteQuantity MOD 256);
    n := cbSrcLength;
    IF n > 242 THEN
        n := 242;
    END_IF;
    mb.DATA[8] := UDINT_TO_BYTE(n);
    i := 0;
    WHILE i < n DO
        mb.DATA[9 + i] := pSrcData[i];
        i := i + 1;
    END_WHILE;
    mb.RLEN := 9 + n;
    mb.EXEC := bExecute;
    mb();
    bBusy := mb.BUSY;
    bDone := mb.DONE;
    IF mb.DONE THEN
        i := 0;
        WHILE i < mb.DLEN AND i < 256 DO
            pDestData[i] := mb.DATA[i];
            i := i + 1;
        END_WHILE;
        cbRead := mb.DLEN;
    END_IF;
    nErrId := mb.ERRID;
    IF mb.RESULT = 1 THEN
        nErrId := 16#8000 + mb.EXC;
    END_IF;
    bError := (mb.ERRID <> 0) OR (mb.RESULT = 1);
END_FUNCTION_BLOCK

FUNCTION_BLOCK FB_MBRtuDiagnose
VAR_INPUT
    sDevice : STRING[63];
    nBaud : UDINT := 9600;
    nParity : UDINT := 0;
    nDataBits : UDINT := 8;
    nStopBits : UDINT := 1;
    nUnitID : BYTE := 1;
    nWriteData : WORD;
    bExecute : BOOL;
    tTimeout : TIME;
END_VAR
VAR_OUTPUT
    bBusy : BOOL;
    bDone : BOOL;
    bError : BOOL;
    nErrId : UDINT;
    cbRead : UDINT;
    pData : ARRAY[0..255] OF BYTE;
END_VAR
VAR
    mb : FB_ModbusRtu;
    i : UDINT;
END_VAR
    mb.FUNC := 8;
    mb.DEV := sDevice;
    mb.BAUD := nBaud;
    mb.PARITY := nParity;
    mb.DBITS := nDataBits;
    mb.SBITS := nStopBits;
    mb.UNIT := nUnitID;
    mb.TIMEOUT := tTimeout;
    mb.DATA[0] := UINT_TO_BYTE(nWriteData / 256);
    mb.DATA[1] := UINT_TO_BYTE(nWriteData MOD 256);
    mb.RLEN := 2;
    mb.EXEC := bExecute;
    mb();
    bBusy := mb.BUSY;
    bDone := mb.DONE;
    IF mb.DONE THEN
        i := 0;
        WHILE i < mb.DLEN AND i < 256 DO
            pData[i] := mb.DATA[i];
            i := i + 1;
        END_WHILE;
        cbRead := mb.DLEN;
    END_IF;
    nErrId := mb.ERRID;
    IF mb.RESULT = 1 THEN
        nErrId := 16#8000 + mb.EXC;
    END_IF;
    bError := (mb.ERRID <> 0) OR (mb.RESULT = 1);
END_FUNCTION_BLOCK
